Staubli VAL3: insertDelay1.pgx

public program insertDelay1()
  local bool l_bExit
  local bool l_bResult
  local num l_nPoint
begin
  do

    //    if util:sPage!="insertDelay"
    //      util:sPage="insertDelay"
    //      nSetDelay=0
    //      userPageBindClick("insertDelay","btn1",bConfirmDelay,true)
    //      userPageBindClick("insertDelay","btn2",bBackDelay,true)
    //      userPageBind("insertDelay","nmb1","value",nSetDelay,1,"rw")
    //      userPage(util:sPage)
    //      delay(0.5)

    //    endIf

    //2024.11.20 add 插入喷淋延时由上位机控制时长s
    //    if bConfirmDelay
    //      bConfirmDelay=false
    nSetDelay=0
    call trajectory:getPointIndex(sTrajItem,sSelPoint,l_nPoint,l_bResult)
    call trajectory:insertDelay(sTrajItem,l_nPoint,bToSave,11,nSetDelay)
    l_bExit=true

    //    elseIf bBackDelay
    //      bBackDelay=false
    //      l_bExit=true
    //    endIf



    delay(0)
  until l_bExit==true
end
